FUNCTION_BLOCK FB_TestableTon
VAR_INPUT
    IN : BOOL;
    PT : TIME;
    TestMode : BOOL;
    TestDone : BOOL;
END_VAR

VAR_OUTPUT
    Q : BOOL;
    ET : TIME;
END_VAR

VAR
    InternalTON : TON;
END_VAR


IF TestMode THEN
    Q := IN AND TestDone;
    ET := T#0MS;
ELSE
    InternalTON(
        IN := IN,
        PT := PT
    );

    Q := InternalTON.Q;
    ET := InternalTON.ET;
END_IF

END_FUNCTION_BLOCK

(* stored: Version 1.1.0.1, ProductVersion 3.1.4024.9
   POU FB_TestableTon: Id {e46f90b1-57b7-4c55-ac15-d319d8bcede7}, SpecialFunc None *)
